(* IEC 61131-3 sources: Caravan/Archiv/12-04-19/Stations/MachineControl/MachineControl/Network/Manage_Net, 1 file *)

(* ---- ONE_Manage_Net_Table.st ---- *)
#define OBJECTS_CONFIG

FUNCTION GLOBAL TAB ONE_Manage_Net
-1$UINT, 0$UINT,
0$UINT, 0$UINT,

1$UDINT,
TO_UDINT(440431991), "Timer_Class", 0$UINT, 0$UINT, 1$UINT,

_NO_ATTR, TO_UDINT(1302809437), "TIMER_CLASS1",

//Internal connections
0$UDINT,
0$UDINT,
0$UDINT,
0$UDINT,

//Initialization values
0$UDINT,
0$UDINT,

//Symbolic initialization values
0$UDINT,
0$UDINT,

//Initialization of string values
0$UDINT,
0$UDINT,

//Configuration of tasks (RealTime, Cyclic, Background)
0$UDINT,
0$UDINT,

0$UDINT,
1$UDINT,
TO_UDINT(0), (-2147483548)$UDINT, 4194303$DINT, 	//TIMER_CLASS1

0$UDINT,
0$UDINT,

//External connections
0$UDINT,
0$UDINT,

//Magic internal connections
0$UDINT,
0$UDINT,

//Configuration of timeslots of tasks (RealTime, Cyclic)
#ifdef __LSLLDR_TIMESLOTS__
0$UDINT,
0$UDINT,

0$UDINT,
0$UDINT,

#endif //__LSLLDR_TIMESLOTS__

//MultiMaster connections
#ifdef __LSLLDR_MULTIMASTER__
0$UDINT,
0$UDINT,
#endif //__LSLLDR_MULTIMASTER__

//Configuration for task ID (RealTime, CyclicTime)
#ifdef __LSLLDR_TASKID__
"\\\\TASKS2  "
0$UDINT,
0$UDINT,

0$UDINT,
1$UDINT,
(0)$UDINT, 	//TIMER_CLASS1

0$UDINT,
0$UDINT,

#endif //__LSLLDR_TASKID__

END_FUNCTION
